// TIA Portal project "FactoryIO_Template_S7-1200_V15_V18_6" (V18)
// Vorlageprojekt für das Buch mit Zielsystem S7-1200

(* hardware
DEVICE "S7-1200-Station_1"  S7-1200 Station
   slot 0: "Baugruppenträger_0"  Rack  V1.0
   slot 1: "PLC_1"  CPU 1214C AC/DC/Rly  6ES7 214-1BG40-0XB0  V4.6
   slot 2: "AI 4xTC_1"  SM 1231 AI4 x TC  6ES7 231-5QD32-0XB0  V2.0
   slot 3: "AQ 4x14BIT_1"  6ES7 232-4HD32-0XB0  V2.1
   slot 4: "AQ 4x14BIT_2"  6ES7 232-4HD32-0XB0  V2.1
*)

// ===== PLC "PLC_1"  CPU 1214C AC/DC/Rly =====

VAR_GLOBAL   // PLC tag table "Standard-Variablentabelle"
   "Sistem Start" AT %I0.0 : Bool;
   "Sistem Stop" AT %I0.1 : Bool;
   "Termokupl Girişi" AT %IW96 : Int;
   "Fan 1" AT %QW30 : Int;
   "Fan 2" AT %QW32 : Int;
   "Fan 3" AT %QW34 : Int;
   "Fan 4" AT %QW40 : Int;
   "Fan 5" AT %QW42 : Int;
   "Fan 6" AT %QW44 : Int;
   "Düşük Sıcaklık Lambası" AT %Q0.0 : Bool;
   "Normal Sıcaklık Lambası" AT %Q0.1 : Bool;
   "Yüksek Sıcaklık Lambası" AT %Q0.2 : Bool;
   "Çok Yüksek Sıcaklık Lambası" AT %Q0.3 : Bool;
   "Tag_1" AT %MW10 : Int;
   "Tag_2" AT %MD12 : Real;
   "Ortam Sıcaklığı" AT %MD16 : Real;
   "System_Byte" AT %MB1 : Byte;
   "FirstScan" AT %M1.0 : Bool;
   "DiagStatusUpdate" AT %M1.1 : Bool;
   "AlwaysTRUE" AT %M1.2 : Bool;
   "AlwaysFALSE" AT %M1.3 : Bool;
   "Clock_Byte" AT %MB0 : Byte;
   "Clock_10Hz" AT %M0.0 : Bool;
   "Clock_5Hz" AT %M0.1 : Bool;
   "Clock_2.5Hz" AT %M0.2 : Bool;
   "Clock_2Hz" AT %M0.3 : Bool;
   "Clock_1.25Hz" AT %M0.4 : Bool;
   "Clock_1Hz" AT %M0.5 : Bool;
   "Clock_0.625Hz" AT %M0.6 : Bool;
   "Clock_0.5Hz" AT %M0.7 : Bool;
   "Çok Yüksek Sıcaklık Mem" AT %M20.0 : Bool;
   "Yüksek Sıcaklık Uyarı Lambası" AT %M20.1 : Bool;
END_VAR

FUNCTION "MHJ-PLC-Lab-Function-S71200" : Void   // FC9000, SCL
{ S7_Optimized_Access := 'TRUE' }
VERSION : 0.1
   VAR_TEMP
      rdTimeReturn : Int;
      outputTime : DTL;
      SyncVal : Byte;
      forVal : Int;
      forVal_2 : Int;
      Value : Byte;
   END_VAR
   VAR CONSTANT
      CompVal : Byte := 16#34;
      Value_01 : Byte := 16#11;
      Value_01_DW : DWord := 16#A165_D992;
      Value_02_DW : DWord := 16#58BE_4401;
   END_VAR
BEGIN

   #Value:=PEEK(area := 16#82,
        dbNumber := 0,
        byteOffset := 511);
   #Value := #Value + 1;

   POKE(area := 16#82,
        dbNumber := 0,
        byteOffset := 511,
        value := #Value);

   POKE(area:=16#81,
        dbNumber:=0,
        byteOffset:=1016,
        value:=#Value_01_DW);
   POKE(area := 16#81,
        dbNumber := 0,
        byteOffset := 1020,
        value := #Value_02_DW);

   POKE(area := 16#81,
        dbNumber := 0,
        byteOffset := 511,
        value := B#16#00);

   FOR #forVal := 0 TO 120 DO
       FOR #forVal_2:=0 TO 10 DO
           #rdTimeReturn:=RD_SYS_T(#outputTime);
           #rdTimeReturn := WR_SYS_T(#outputTime);
           #rdTimeReturn := RD_SYS_T(#outputTime);
           #rdTimeReturn := WR_SYS_T(#outputTime);
       END_FOR;
       #SyncVal:= PEEK(area := 16#81,
                      dbNumber := 0,
                      byteOffset := 511);
       IF #SyncVal = #CompVal THEN
          GOTO M_1;
       END_IF;
   END_FOR;
   RETURN;

   M_1:
   POKE(area := 16#81,
        dbNumber := 0,
        byteOffset := 511,
        value := B#16#0);
END_FUNCTION

ORGANIZATION_BLOCK "Main"   // OB1, LAD, ProgramCycle
TITLE = "Main Program Sweep (Cycle)"
{ S7_Optimized_Access := 'TRUE' }
VERSION : 0.1
   VAR_INPUT
      Initial_Call : Bool;   // Initial call of this OB
      Remanence : Bool;   // =True, if remanent data are available
   END_VAR
   VAR_TEMP   // added for the SCL form of the ladder/FBD networks
      _w1 : Bool;
   END_VAR
BEGIN

REGION Network 1: Konnektierungsbaustein für PLC-Lab / PLC LAB FONKSİYONUNUN ÇAĞRILMASI
   // Im Netzwerk 1 wird der Konnektierungsbaustein für PLC-Lab aufgerufen.
   // Dieser Aufruf darf nicht entfernt werden!
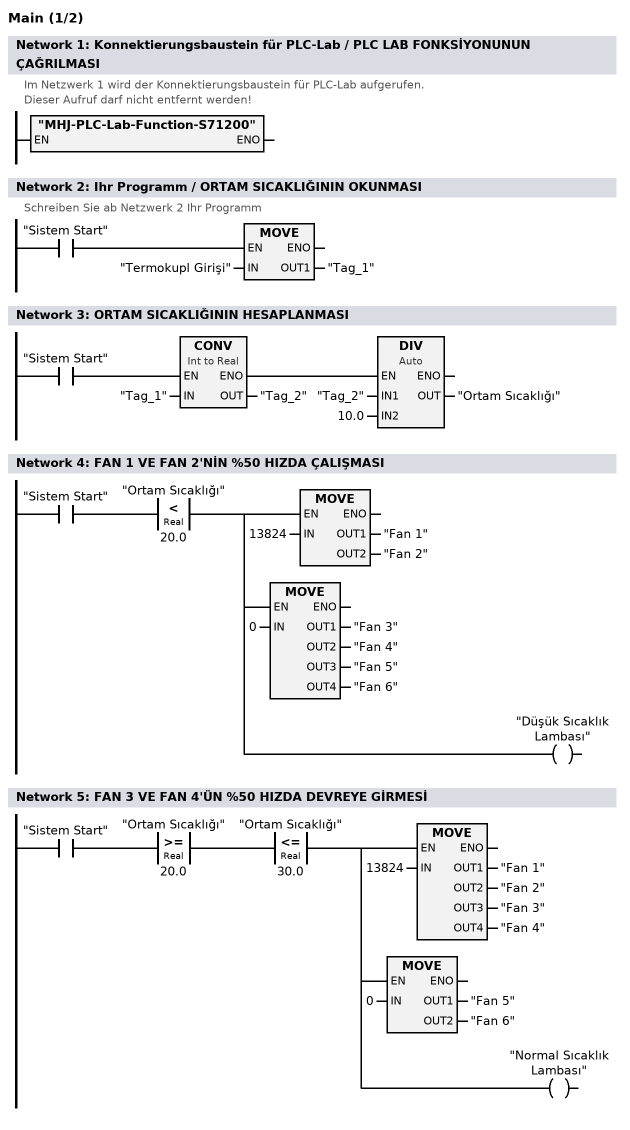
   RUNG wire#powerrail
      "MHJ-PLC-Lab-Function-S71200"()
   END_RUNG
   // the same network as SCL:
   "MHJ-PLC-Lab-Function-S71200"();
END_REGION

REGION Network 2: Ihr Programm / ORTAM SICAKLIĞININ OKUNMASI
   // Schreiben Sie ab Netzwerk 2 Ihr Programm
   RUNG wire#powerrail
      Contact( "Sistem Start" )
      Move(in := "Termokupl Girişi", out1 => "Tag_1")
   END_RUNG
   // the same network as SCL:
   IF "Sistem Start" THEN "Tag_1" := "Termokupl Girişi"; END_IF;
END_REGION

REGION Network 3: ORTAM SICAKLIĞININ HESAPLANMASI
   RUNG wire#powerrail
      Contact( "Sistem Start" )
      { S7_Templates := "[SrcType := Int, DestType := Real]" } Convert(in := "Tag_1", out => "Tag_2")
      Div(in1 := "Tag_2", in2 := 10.0, out => "Ortam Sıcaklığı")
   END_RUNG
   // the same network as SCL:
   IF "Sistem Start" THEN
       "Tag_2" := INT_TO_REAL("Tag_1");
       "Ortam Sıcaklığı" := "Tag_2" / 10.0;
   END_IF;
END_REGION

REGION Network 4: FAN 1 VE FAN 2'NİN %50 HIZDA ÇALIŞMASI
   RUNG wire#powerrail
      Contact( "Sistem Start" )
      { S7_Templates := "SrcType := Real" } LT_Contact(in1 := "Ortam Sıcaklığı", in2 := 20.0)
      wire#w1
      Move(in := 13824, out1 => "Fan 1", out2 => "Fan 2")
   END_RUNG
   RUNG wire#w1
      Move(in := 0, out1 => "Fan 3", out2 => "Fan 4", out3 => "Fan 5", out4 => "Fan 6")
   END_RUNG
   RUNG wire#w1
      Coil( "Düşük Sıcaklık Lambası" )
   END_RUNG
   // the same network as SCL:
   #_w1 := "Sistem Start" AND ("Ortam Sıcaklığı" < 20.0);
   IF #_w1 THEN
       "Fan 1" := 13824;
       "Fan 2" := 13824;
       "Fan 3" := 0;
       "Fan 4" := 0;
       "Fan 5" := 0;
       "Fan 6" := 0;
   END_IF;
   "Düşük Sıcaklık Lambası" := #_w1;
END_REGION

REGION Network 5: FAN 3 VE FAN 4'ÜN %50 HIZDA DEVREYE GİRMESİ
   RUNG wire#powerrail
      Contact( "Sistem Start" )
      { S7_Templates := "SrcType := Real" } GE_Contact(in1 := "Ortam Sıcaklığı", in2 := 20.0)
      { S7_Templates := "SrcType := Real" } LE_Contact(in1 := "Ortam Sıcaklığı", in2 := 30.0)
      wire#w1
      Move(in := 13824, out1 => "Fan 1", out2 => "Fan 2", out3 => "Fan 3", out4 => "Fan 4")
   END_RUNG
   RUNG wire#w1
      Move(in := 0, out1 => "Fan 5", out2 => "Fan 6")
   END_RUNG
   RUNG wire#w1
      Coil( "Normal Sıcaklık Lambası" )
   END_RUNG
   // the same network as SCL:
   #_w1 := "Sistem Start" AND ("Ortam Sıcaklığı" >= 20.0) AND ("Ortam Sıcaklığı" <= 30.0);
   IF #_w1 THEN
       "Fan 1" := 13824;
       "Fan 2" := 13824;
       "Fan 3" := 13824;
       "Fan 4" := 13824;
       "Fan 5" := 0;
       "Fan 6" := 0;
   END_IF;
   "Normal Sıcaklık Lambası" := #_w1;
END_REGION

REGION Network 6: FAN 5 VE FAN 6 CALISMA YUZDE 50
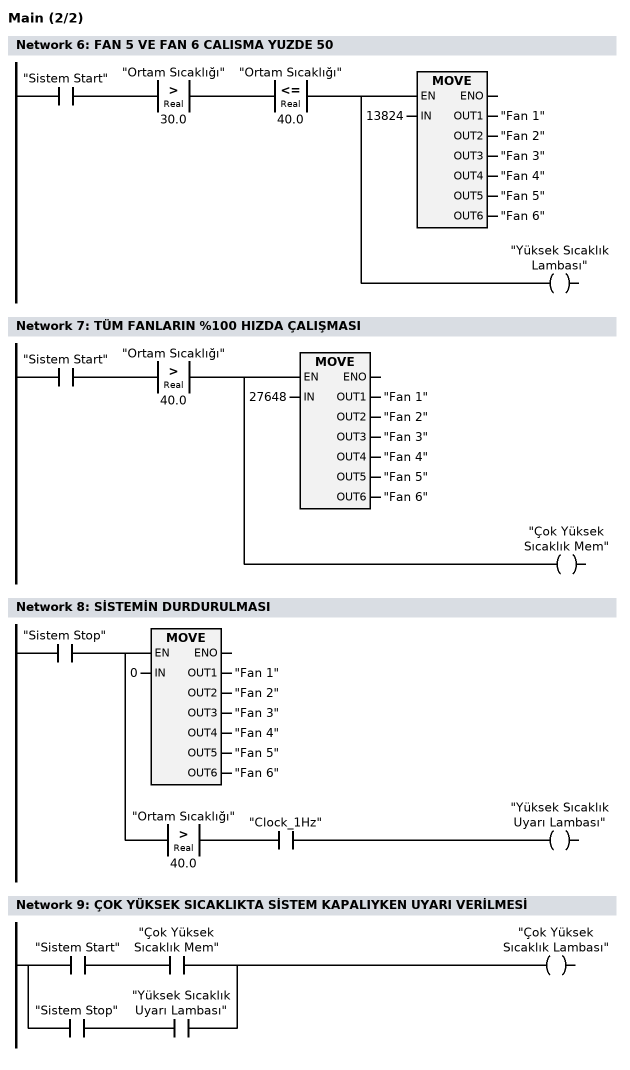
   RUNG wire#powerrail
      Contact( "Sistem Start" )
      { S7_Templates := "SrcType := Real" } GT_Contact(in1 := "Ortam Sıcaklığı", in2 := 30.0)
      { S7_Templates := "SrcType := Real" } LE_Contact(in1 := "Ortam Sıcaklığı", in2 := 40.0)
      wire#w1
      Move(in := 13824, out1 => "Fan 1", out2 => "Fan 2", out3 => "Fan 3", out4 => "Fan 4", out5 => "Fan 5", out6 => "Fan 6")
   END_RUNG
   RUNG wire#w1
      Coil( "Yüksek Sıcaklık Lambası" )
   END_RUNG
   // the same network as SCL:
   #_w1 := "Sistem Start" AND ("Ortam Sıcaklığı" > 30.0) AND ("Ortam Sıcaklığı" <= 40.0);
   IF #_w1 THEN
       "Fan 1" := 13824;
       "Fan 2" := 13824;
       "Fan 3" := 13824;
       "Fan 4" := 13824;
       "Fan 5" := 13824;
       "Fan 6" := 13824;
   END_IF;
   "Yüksek Sıcaklık Lambası" := #_w1;
END_REGION

REGION Network 7: TÜM FANLARIN %100 HIZDA ÇALIŞMASI
   RUNG wire#powerrail
      Contact( "Sistem Start" )
      { S7_Templates := "SrcType := Real" } GT_Contact(in1 := "Ortam Sıcaklığı", in2 := 40.0)
      wire#w1
      Move(in := 27648, out1 => "Fan 1", out2 => "Fan 2", out3 => "Fan 3", out4 => "Fan 4", out5 => "Fan 5", out6 => "Fan 6")
   END_RUNG
   RUNG wire#w1
      Coil( "Çok Yüksek Sıcaklık Mem" )
   END_RUNG
   // the same network as SCL:
   #_w1 := "Sistem Start" AND ("Ortam Sıcaklığı" > 40.0);
   IF #_w1 THEN
       "Fan 1" := 27648;
       "Fan 2" := 27648;
       "Fan 3" := 27648;
       "Fan 4" := 27648;
       "Fan 5" := 27648;
       "Fan 6" := 27648;
   END_IF;
   "Çok Yüksek Sıcaklık Mem" := #_w1;
END_REGION

REGION Network 8: SİSTEMİN DURDURULMASI
   RUNG wire#powerrail
      Contact( "Sistem Stop" )
      wire#w1
      Move(in := 0, out1 => "Fan 1", out2 => "Fan 2", out3 => "Fan 3", out4 => "Fan 4", out5 => "Fan 5", out6 => "Fan 6")
   END_RUNG
   RUNG wire#w1
      { S7_Templates := "SrcType := Real" } GT_Contact(in1 := "Ortam Sıcaklığı", in2 := 40.0)
      Contact( "Clock_1Hz" )
      Coil( "Yüksek Sıcaklık Uyarı Lambası" )
   END_RUNG
   // the same network as SCL:
   IF "Sistem Stop" THEN
       "Fan 1" := 0;
       "Fan 2" := 0;
       "Fan 3" := 0;
       "Fan 4" := 0;
       "Fan 5" := 0;
       "Fan 6" := 0;
   END_IF;
   "Yüksek Sıcaklık Uyarı Lambası" := "Sistem Stop" AND ("Ortam Sıcaklığı" > 40.0) AND "Clock_1Hz";
END_REGION

REGION Network 9: ÇOK YÜKSEK SICAKLIKTA SİSTEM KAPALIYKEN UYARI VERİLMESİ
   RUNG wire#powerrail
      Contact( "Sistem Start" )
      Contact( "Çok Yüksek Sıcaklık Mem" )
      wire#w1
      Coil( "Çok Yüksek Sıcaklık Lambası" )
   END_RUNG
   RUNG wire#powerrail
      Contact( "Sistem Stop" )
      Contact( "Yüksek Sıcaklık Uyarı Lambası" )
   END_RUNG wire#w1
   // the same network as SCL:
   "Çok Yüksek Sıcaklık Lambası" := ("Sistem Start" AND "Çok Yüksek Sıcaklık Mem") OR ("Sistem Stop" AND "Yüksek Sıcaklık Uyarı Lambası");
END_REGION
END_ORGANIZATION_BLOCK